Fanuc KAREL source: ko00063.KL

-- PROVISIONAL review KL for V770-1; original PC SHA256 feabbbcedf3b245b340952a0a87633217282b26df9160add677d54192c530a83
-- Incomplete behavior may be omitted. Consult companion uncertainty JSON. Do not deploy.
PROGRAM KO00063
%NOLOCKGROUP
BEGIN
  -- UNRESOLVED_PC offsets 5-12; opcodes 9D,23
  -- UNRESOLVED_PC offsets 17-69; opcodes 27,27,49,7E,AD,27,49,7E,AD,22,31,7E,4A
  -- UNRESOLVED_PC offsets 74-78; opcodes 7F
END KO00063
